SYSTEM StopperingModule (* Module Stoppering, generated from its module specification *)
  (* Standard: 61499-2 *)
  APPLICATION Stoppering (* Module Stoppering on target pc (localhost, IO modbus; generated by modgen) *)
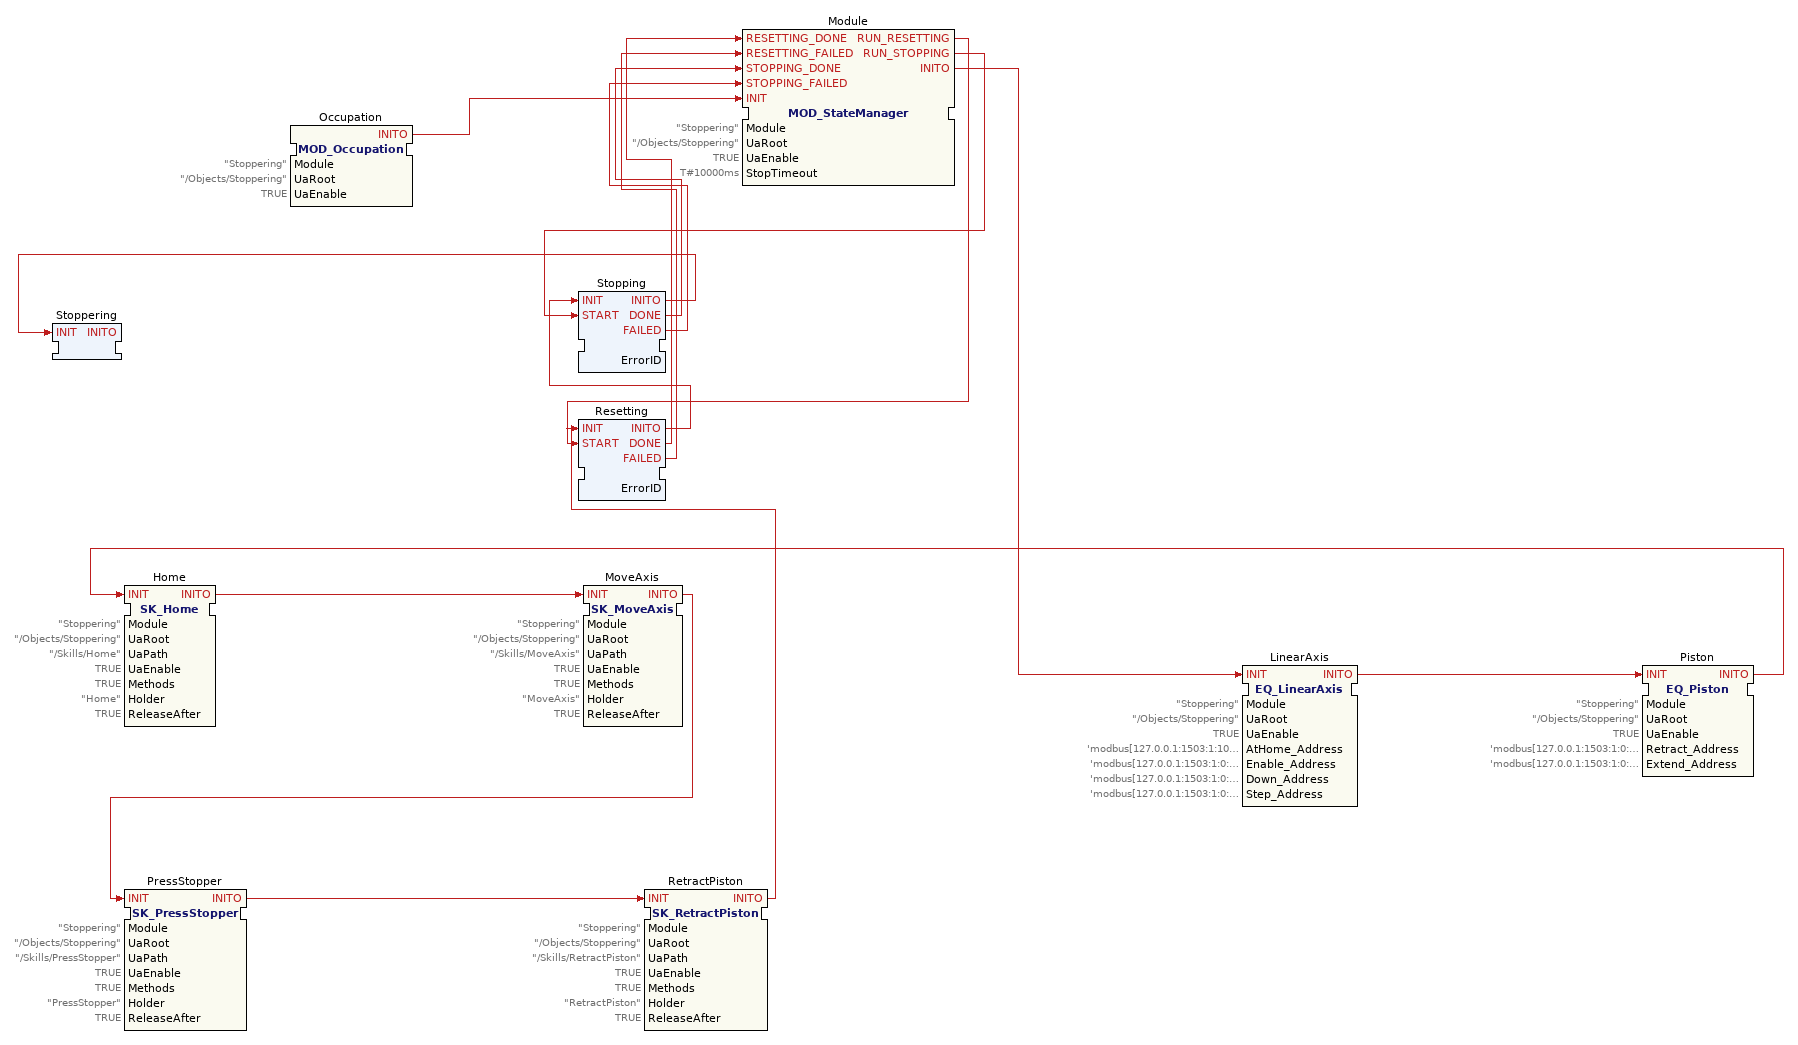
    (* Group ModuleLevel: Module level: occupation, PackML state manager, start-up and the target's IO lines *)
    (* Group ModuleLevelSkills: Module level skills: Control, Sequences (Execute, Stop) of skill primitives and Release; OPC UA /Skills/<name> *)
    (* Group Procedures: Procedures the module state manager runs while Resetting and Stopping *)
    (* Group SkillPrimitives: Skill primitives: one equipment command until a sensor or a time; OPC UA /Skills/<name> *)
    (* Group EquipmentIO: Equipment IO: the only owners of the IO points; skills send them output values over local channels *)
    FBS
      Occupation : modlib::MOD_Occupation(Module := "Stoppering", UaRoot := "/Objects/Stoppering", UaEnable := TRUE); (* Who may command the module. A client calls Occupy(Session) at /Objects/Stoppering/Occupation first; until it calls Release, only commands with that session id are accepted. Every block hears the owner on loc[Stoppering/owner]. *) {SET_ATTRIBUTE(GroupName, ModuleLevel)}
      Module : modlib::MOD_StateManager(Module := "Stoppering", UaRoot := "/Objects/Stoppering", UaEnable := TRUE, StopTimeout := T#10000ms); (* The module's PackML state. The owner calls Reset, Start, Stop, Abort or Clear at /Objects/Stoppering/Module; State is at /Objects/Stoppering/Module/State and on loc[Stoppering/state]. Reset runs the Resetting procedure, Stop the Stopping procedure; skills may be started only in Execute. *) {SET_ATTRIBUTE(GroupName, ModuleLevel)}
      LinearAxis : stoppering::EQ_LinearAxis(Module := "Stoppering", UaRoot := "/Objects/Stoppering", UaEnable := TRUE, AtHome_Address := 'modbus[127.0.0.1:1503:1:10:d0:]', Enable_Address := 'modbus[127.0.0.1:1503:1:0::c0]', Down_Address := 'modbus[127.0.0.1:1503:1:0::c1]', Step_Address := 'modbus[127.0.0.1:1503:1:0::h0]'); (* Equipment LinearAxis: Lift of the stoppering head, a stepper motor through a step and direction driver, with a limit switch at the top (home). The only block that touches its pins (AtHome = modbus[127.0.0.1:1503:1:10:d0:], Enable = modbus[127.0.0.1:1503:1:0::c0], Down = modbus[127.0.0.1:1503:1:0::c1], Step = modbus[127.0.0.1:1503:1:0::h0]). Skills send it what to switch on loc[Stoppering/LinearAxis/cmd]; it reports its inputs on loc[Stoppering/LinearAxis/state] and at /Objects/Stoppering/Equipment/LinearAxis. *) {SET_ATTRIBUTE(GroupName, EquipmentIO)}
      Piston : stoppering::EQ_Piston(Module := "Stoppering", UaRoot := "/Objects/Stoppering", UaEnable := TRUE, Retract_Address := 'modbus[127.0.0.1:1503:1:0::c2]', Extend_Address := 'modbus[127.0.0.1:1503:1:0::c3]'); (* Equipment Piston: Small linear actuator that presses the stopper in, through an L298N (IN1 retract, IN2 extend); no sensors. The only block that touches its pins (Retract = modbus[127.0.0.1:1503:1:0::c2], Extend = modbus[127.0.0.1:1503:1:0::c3]). Skills send it what to switch on loc[Stoppering/Piston/cmd]; it reports its inputs on loc[Stoppering/Piston/state] and at /Objects/Stoppering/Equipment/Piston. *) {SET_ATTRIBUTE(GroupName, EquipmentIO)}
      Home : stoppering::SK_Home(Module := "Stoppering", UaRoot := "/Objects/Stoppering", UaPath := "/Skills/Home", UaEnable := TRUE, Methods := TRUE, Holder := "Home", ReleaseAfter := TRUE); (* Skill Home, offered on its own: Head up to the limit switch; from there its position is known, using LinearAxis. A client calls Start (with the parameters), Stop, Abort or Reset at /Objects/Stoppering/Skills/Home; State, ErrorID, Parameters and Results are there too. *) {SET_ATTRIBUTE(GroupName, SkillPrimitives)}
      MoveAxis : stoppering::SK_MoveAxis(Module := "Stoppering", UaRoot := "/Objects/Stoppering", UaPath := "/Skills/MoveAxis", UaEnable := TRUE, Methods := TRUE, Holder := "MoveAxis", ReleaseAfter := TRUE); (* Skill MoveAxis, offered on its own: Head to Position, measured down from the limit switch; the direction follows from where it is, using LinearAxis. A client calls Start (with the parameters), Stop, Abort or Reset at /Objects/Stoppering/Skills/MoveAxis; State, ErrorID, Parameters and Results are there too. *) {SET_ATTRIBUTE(GroupName, SkillPrimitives)}
      PressStopper : stoppering::SK_PressStopper(Module := "Stoppering", UaRoot := "/Objects/Stoppering", UaPath := "/Skills/PressStopper", UaEnable := TRUE, Methods := TRUE, Holder := "PressStopper", ReleaseAfter := TRUE); (* Skill PressStopper, offered on its own: Press the stopper in, the piston out for the stroke and back in (open loop, by time), using Piston. A client calls Start (with the parameters), Stop, Abort or Reset at /Objects/Stoppering/Skills/PressStopper; State, ErrorID, Parameters and Results are there too. *) {SET_ATTRIBUTE(GroupName, SkillPrimitives)}
      RetractPiston : stoppering::SK_RetractPiston(Module := "Stoppering", UaRoot := "/Objects/Stoppering", UaPath := "/Skills/RetractPiston", UaEnable := TRUE, Methods := TRUE, Holder := "RetractPiston", ReleaseAfter := TRUE); (* Skill RetractPiston, offered on its own: Piston back in for the stroke (open loop); for a piston left out by an abort, using Piston. A client calls Start (with the parameters), Stop, Abort or Reset at /Objects/Stoppering/Skills/RetractPiston; State, ErrorID, Parameters and Results are there too. *) {SET_ATTRIBUTE(GroupName, SkillPrimitives)}
    END_FBS
    SUBAPPLICATION Resetting (* Procedure the module runs while Resetting *)
      {SET_ATTRIBUTE(GroupName, Procedures)}
      EVENT_INPUT
        INIT : EInit;
        START;
      END_EVENT
      EVENT_OUTPUT
        INITO : EInit;
        DONE;
        FAILED;
      END_EVENT
      VAR_OUTPUT
        ErrorID : UINT;
      END_VAR
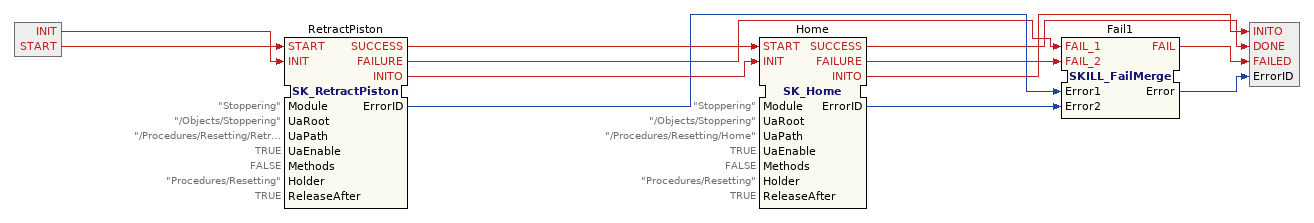
      FBS
        RetractPiston : stoppering::SK_RetractPiston(Module := "Stoppering", UaRoot := "/Objects/Stoppering", UaPath := "/Procedures/Resetting/RetractPiston", UaEnable := TRUE, Methods := FALSE, Holder := "Procedures/Resetting", ReleaseAfter := TRUE); (* Step 1 of Resetting: runs the skill RetractPiston. Its State and ErrorID are at /Objects/Stoppering/Procedures/Resetting/RetractPiston; it keeps the equipment under the name Procedures/Resetting. *)
        Home : stoppering::SK_Home(Module := "Stoppering", UaRoot := "/Objects/Stoppering", UaPath := "/Procedures/Resetting/Home", UaEnable := TRUE, Methods := FALSE, Holder := "Procedures/Resetting", ReleaseAfter := TRUE); (* Step 2 of Resetting: runs the skill Home. Its State and ErrorID are at /Objects/Stoppering/Procedures/Resetting/Home; it keeps the equipment under the name Procedures/Resetting. *)
        Fail1 : modlib::SKILL_FailMerge; (* Joins the failures of the steps into one (with its error code), so any step's failure ends the sequence. *)
      END_FBS
      EVENT_CONNECTIONS
        RetractPiston.SUCCESS TO Home.START;
        START TO RetractPiston.START;
        Home.SUCCESS TO DONE;
        RetractPiston.FAILURE TO Fail1.FAIL_1;
        Home.FAILURE TO Fail1.FAIL_2;
        Fail1.FAIL TO FAILED;
        INIT TO RetractPiston.INIT;
        Home.INITO TO INITO;
        RetractPiston.INITO TO Home.INIT;
      END_CONNECTIONS
      DATA_CONNECTIONS
        RetractPiston.ErrorID TO Fail1.Error1;
        Home.ErrorID TO Fail1.Error2;
        Fail1.Error TO ErrorID;
      END_CONNECTIONS
    END_SUBAPPLICATION
    SUBAPPLICATION Stopping (* Procedure the module runs while Stopping *)
      {SET_ATTRIBUTE(GroupName, Procedures)}
      EVENT_INPUT
        INIT : EInit;
        START;
      END_EVENT
      EVENT_OUTPUT
        INITO : EInit;
        DONE;
        FAILED;
      END_EVENT
      VAR_OUTPUT
        ErrorID : UINT;
      END_VAR
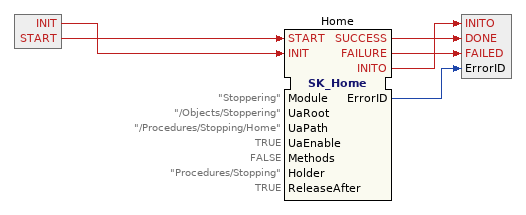
      FBS
        Home : stoppering::SK_Home(Module := "Stoppering", UaRoot := "/Objects/Stoppering", UaPath := "/Procedures/Stopping/Home", UaEnable := TRUE, Methods := FALSE, Holder := "Procedures/Stopping", ReleaseAfter := TRUE); (* Step 1 of Stopping: runs the skill Home. Its State and ErrorID are at /Objects/Stoppering/Procedures/Stopping/Home; it keeps the equipment under the name Procedures/Stopping. *)
      END_FBS
      EVENT_CONNECTIONS
        START TO Home.START;
        Home.SUCCESS TO DONE;
        Home.FAILURE TO FAILED;
        INIT TO Home.INIT;
        Home.INITO TO INITO;
      END_CONNECTIONS
      DATA_CONNECTIONS
        Home.ErrorID TO ErrorID;
      END_CONNECTIONS
    END_SUBAPPLICATION
    SUBAPPLICATION Stoppering (* Module level skill Stoppering: Head down onto the vial, press the stopper in, head up again *)
      {SET_ATTRIBUTE(GroupName, ModuleLevelSkills)}
      EVENT_INPUT
        INIT : EInit;
      END_EVENT
      EVENT_OUTPUT
        INITO : EInit;
      END_EVENT
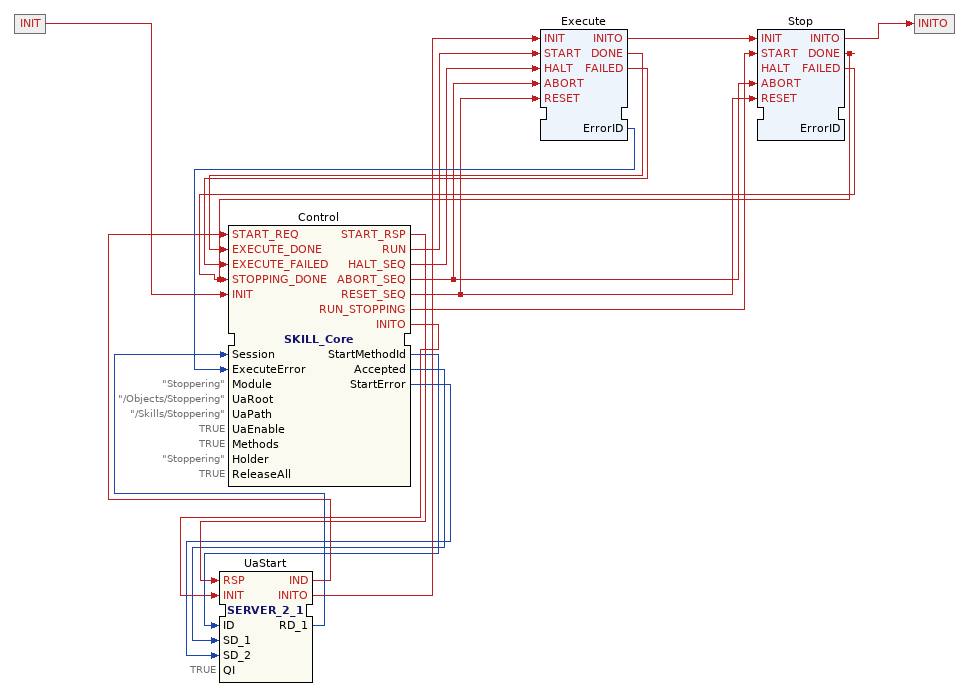
      (* Group Core: The skill's state machine: Stop, Abort, Reset, State and ErrorID over OPC UA; gives up everything the skill holds when a run ends *)
      (* Group Start: The Start method: one block per parameter (range check, value for this run), the values published *)
      (* Group Sequences: What the skill does: Execute, and Stop when it is interrupted; private skill primitives in order *)
      FBS
        Control : modlib::SKILL_Core(Module := "Stoppering", UaRoot := "/Objects/Stoppering", UaPath := "/Skills/Stoppering", UaEnable := TRUE, Methods := TRUE, Holder := "Stoppering", ReleaseAll := TRUE); (* The state machine of the skill Stoppering: checks a client's Start (occupation, module in Execute, not running, values in range), publishes State and ErrorID at /Objects/Stoppering/Skills/Stoppering, offers Stop, Abort and Reset there, starts Execute and runs Stop when the skill is stopped. *) {SET_ATTRIBUTE(GroupName, Core)}
        UaStart : iec61499::net::SERVER_2_1(QI := TRUE); (* The OPC UA method Start of Stoppering: a client's call (session id and parameters) arrives here; the parameters are checked, then Control answers Accepted or an error code. *) {SET_ATTRIBUTE(GroupName, Start)}
      END_FBS
      SUBAPPLICATION Execute (* Stoppering: execute sequence *)
        {SET_ATTRIBUTE(GroupName, Sequences)}
        EVENT_INPUT
          INIT : EInit;
          START;
          HALT;
          ABORT;
          RESET;
        END_EVENT
        EVENT_OUTPUT
          INITO : EInit;
          DONE;
          FAILED;
        END_EVENT
        VAR_OUTPUT
          ErrorID : UINT;
        END_VAR
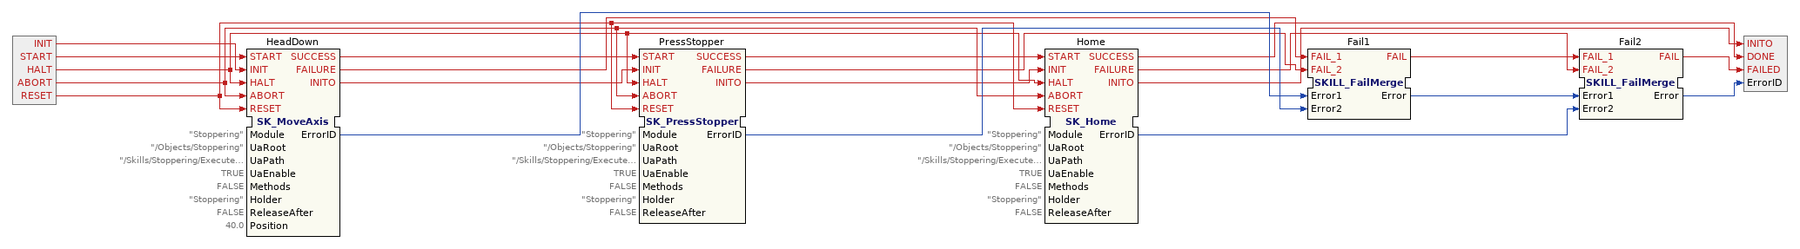
        FBS
          HeadDown : stoppering::SK_MoveAxis(Module := "Stoppering", UaRoot := "/Objects/Stoppering", UaPath := "/Skills/Stoppering/Execute/HeadDown", UaEnable := TRUE, Methods := FALSE, Holder := "Stoppering", ReleaseAfter := FALSE, Position := 40.0); (* Step 1 of Stoppering / Execute: runs the skill MoveAxis with Position = 40.0. Its State and ErrorID are at /Objects/Stoppering/Skills/Stoppering/Execute/HeadDown; it keeps the equipment under the name Stoppering. *)
          PressStopper : stoppering::SK_PressStopper(Module := "Stoppering", UaRoot := "/Objects/Stoppering", UaPath := "/Skills/Stoppering/Execute/PressStopper", UaEnable := TRUE, Methods := FALSE, Holder := "Stoppering", ReleaseAfter := FALSE); (* Step 2 of Stoppering / Execute: runs the skill PressStopper. Its State and ErrorID are at /Objects/Stoppering/Skills/Stoppering/Execute/PressStopper; it keeps the equipment under the name Stoppering. *)
          Home : stoppering::SK_Home(Module := "Stoppering", UaRoot := "/Objects/Stoppering", UaPath := "/Skills/Stoppering/Execute/Home", UaEnable := TRUE, Methods := FALSE, Holder := "Stoppering", ReleaseAfter := FALSE); (* Step 3 of Stoppering / Execute: runs the skill Home. Its State and ErrorID are at /Objects/Stoppering/Skills/Stoppering/Execute/Home; it keeps the equipment under the name Stoppering. *)
          Fail1 : modlib::SKILL_FailMerge; (* Joins the failures of the steps into one (with its error code), so any step's failure ends the sequence. *)
          Fail2 : modlib::SKILL_FailMerge; (* Joins the failures of the steps into one (with its error code), so any step's failure ends the sequence. *)
        END_FBS
        EVENT_CONNECTIONS
          HeadDown.SUCCESS TO PressStopper.START;
          PressStopper.SUCCESS TO Home.START;
          START TO HeadDown.START;
          Home.SUCCESS TO DONE;
          HeadDown.FAILURE TO Fail1.FAIL_1;
          PressStopper.FAILURE TO Fail1.FAIL_2;
          Fail1.FAIL TO Fail2.FAIL_1;
          Home.FAILURE TO Fail2.FAIL_2;
          Fail2.FAIL TO FAILED;
          INIT TO HeadDown.INIT;
          Home.INITO TO INITO;
          HeadDown.INITO TO PressStopper.INIT;
          PressStopper.INITO TO Home.INIT;
          HALT TO HeadDown.HALT;
          HALT TO PressStopper.HALT;
          HALT TO Home.HALT;
          ABORT TO HeadDown.ABORT;
          ABORT TO PressStopper.ABORT;
          ABORT TO Home.ABORT;
          RESET TO HeadDown.RESET;
          RESET TO PressStopper.RESET;
          RESET TO Home.RESET;
        END_CONNECTIONS
        DATA_CONNECTIONS
          HeadDown.ErrorID TO Fail1.Error1;
          PressStopper.ErrorID TO Fail1.Error2;
          Fail1.Error TO Fail2.Error1;
          Home.ErrorID TO Fail2.Error2;
          Fail2.Error TO ErrorID;
        END_CONNECTIONS
      END_SUBAPPLICATION
      SUBAPPLICATION Stop (* Stoppering: stop sequence *)
        {SET_ATTRIBUTE(GroupName, Sequences)}
        EVENT_INPUT
          INIT : EInit;
          START;
          HALT;
          ABORT;
          RESET;
        END_EVENT
        EVENT_OUTPUT
          INITO : EInit;
          DONE;
          FAILED;
        END_EVENT
        VAR_OUTPUT
          ErrorID : UINT;
        END_VAR
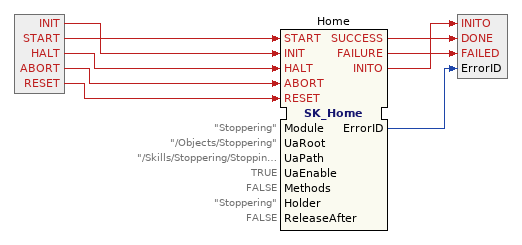
        FBS
          Home : stoppering::SK_Home(Module := "Stoppering", UaRoot := "/Objects/Stoppering", UaPath := "/Skills/Stoppering/Stopping/Home", UaEnable := TRUE, Methods := FALSE, Holder := "Stoppering", ReleaseAfter := FALSE); (* Step 1 of Stoppering / Stop: runs the skill Home. Its State and ErrorID are at /Objects/Stoppering/Skills/Stoppering/Stopping/Home; it keeps the equipment under the name Stoppering. *)
        END_FBS
        EVENT_CONNECTIONS
          START TO Home.START;
          Home.SUCCESS TO DONE;
          Home.FAILURE TO FAILED;
          INIT TO Home.INIT;
          Home.INITO TO INITO;
          HALT TO Home.HALT;
          ABORT TO Home.ABORT;
          RESET TO Home.RESET;
        END_CONNECTIONS
        DATA_CONNECTIONS
          Home.ErrorID TO ErrorID;
        END_CONNECTIONS
      END_SUBAPPLICATION
      EVENT_CONNECTIONS
        Control.START_RSP TO UaStart.RSP;
        UaStart.IND TO Control.START_REQ;
        Control.RUN TO Execute.START;
        Control.HALT_SEQ TO Execute.HALT;
        Control.ABORT_SEQ TO Execute.ABORT;
        Control.RESET_SEQ TO Execute.RESET;
        Execute.DONE TO Control.EXECUTE_DONE;
        Execute.FAILED TO Control.EXECUTE_FAILED;
        Control.RUN_STOPPING TO Stop.START;
        Control.ABORT_SEQ TO Stop.ABORT;
        Control.RESET_SEQ TO Stop.RESET;
        Stop.DONE TO Control.STOPPING_DONE;
        Stop.FAILED TO Control.STOPPING_DONE;
        INIT TO Control.INIT;
        Control.INITO TO UaStart.INIT;
        UaStart.INITO TO Execute.INIT;
        Execute.INITO TO Stop.INIT;
        Stop.INITO TO INITO;
      END_CONNECTIONS
      DATA_CONNECTIONS
        Control.StartMethodId TO UaStart.ID;
        UaStart.RD_1 TO Control.Session;
        Control.Accepted TO UaStart.SD_1;
        Control.StartError TO UaStart.SD_2;
        Execute.ErrorID TO Control.ExecuteError;
      END_CONNECTIONS
    END_SUBAPPLICATION
    EVENT_CONNECTIONS
      Module.RUN_RESETTING TO Resetting.START;
      Resetting.DONE TO Module.RESETTING_DONE;
      Resetting.FAILED TO Module.RESETTING_FAILED;
      Module.RUN_STOPPING TO Stopping.START;
      Stopping.DONE TO Module.STOPPING_DONE;
      Stopping.FAILED TO Module.STOPPING_FAILED;
      Occupation.INITO TO Module.INIT;
      Module.INITO TO LinearAxis.INIT;
      LinearAxis.INITO TO Piston.INIT;
      Piston.INITO TO Home.INIT;
      Home.INITO TO MoveAxis.INIT;
      MoveAxis.INITO TO PressStopper.INIT;
      PressStopper.INITO TO RetractPiston.INIT;
      RetractPiston.INITO TO Resetting.INIT;
      Resetting.INITO TO Stopping.INIT;
      Stopping.INITO TO Stoppering.INIT;
    END_CONNECTIONS
  END_APPLICATION
  APPLICATION Stoppering_pi (* Module Stoppering on target pi (192.168.0.134, IO gpio; generated by modgen) *)
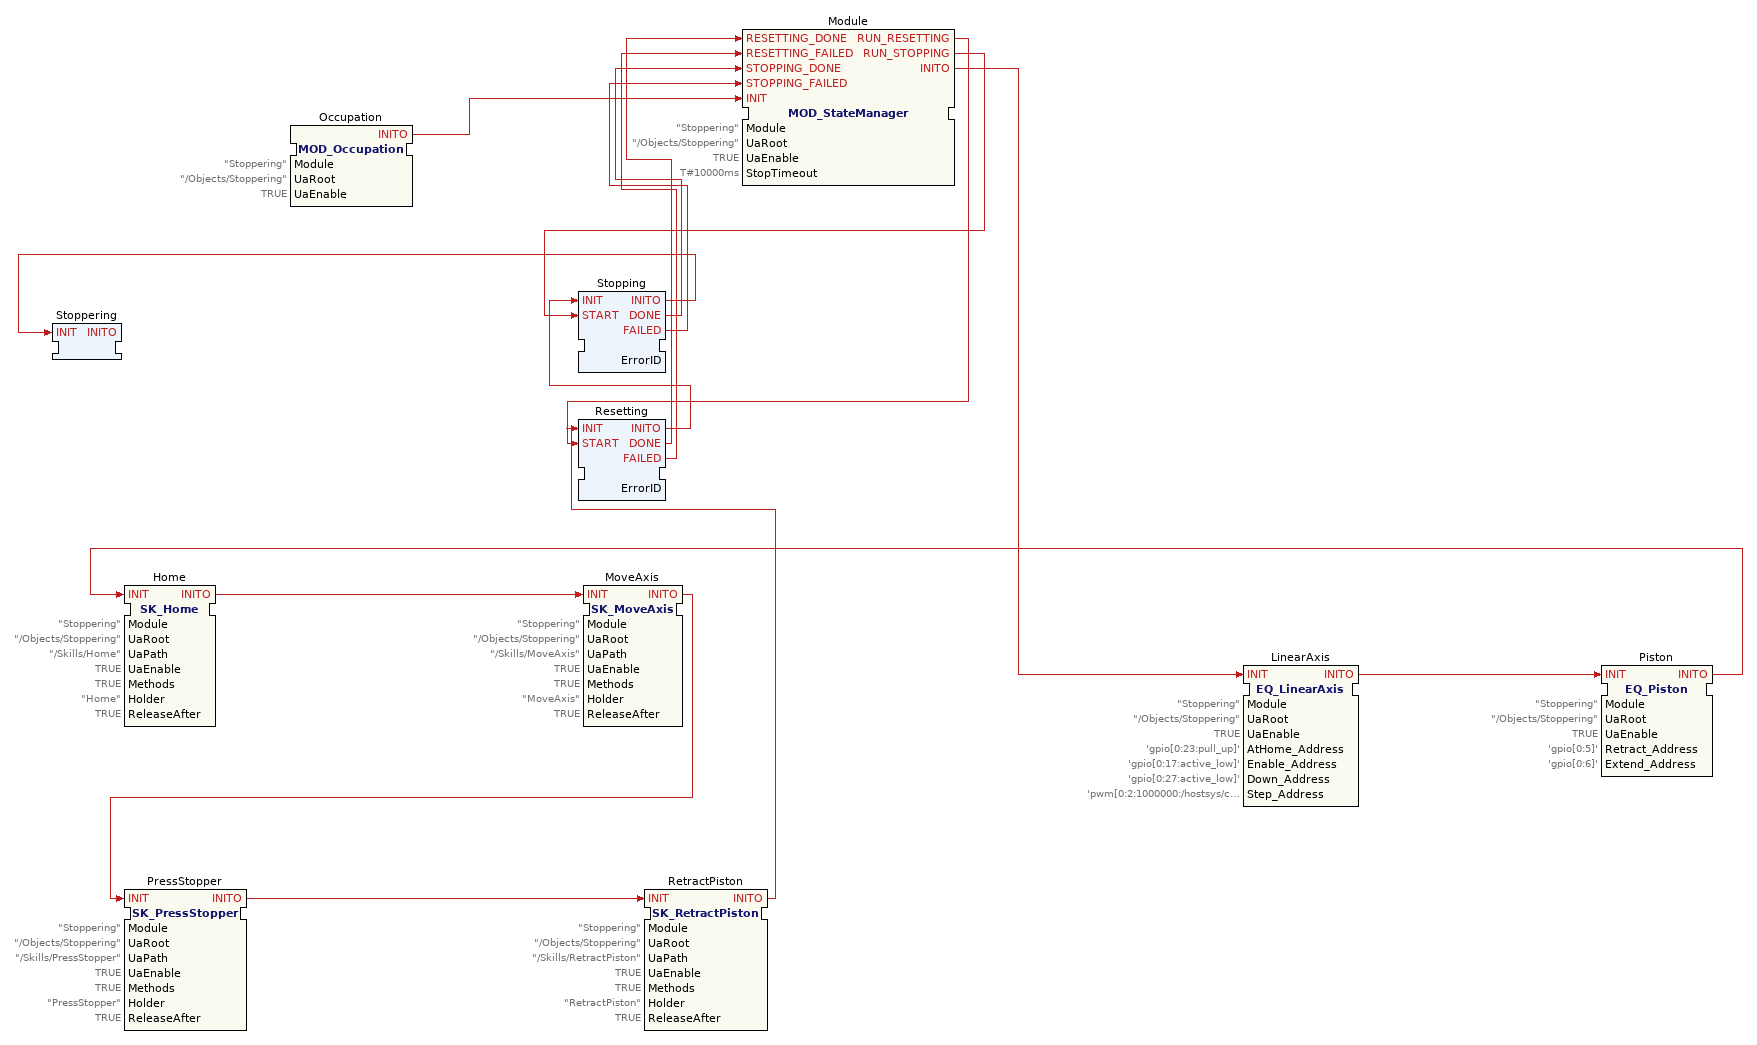
    (* Group ModuleLevel: Module level: occupation, PackML state manager, start-up and the target's IO lines *)
    (* Group ModuleLevelSkills: Module level skills: Control, Sequences (Execute, Stop) of skill primitives and Release; OPC UA /Skills/<name> *)
    (* Group Procedures: Procedures the module state manager runs while Resetting and Stopping *)
    (* Group SkillPrimitives: Skill primitives: one equipment command until a sensor or a time; OPC UA /Skills/<name> *)
    (* Group EquipmentIO: Equipment IO: the only owners of the IO points; skills send them output values over local channels *)
    FBS
      Occupation : modlib::MOD_Occupation(Module := "Stoppering", UaRoot := "/Objects/Stoppering", UaEnable := TRUE); (* Who may command the module. A client calls Occupy(Session) at /Objects/Stoppering/Occupation first; until it calls Release, only commands with that session id are accepted. Every block hears the owner on loc[Stoppering/owner]. *) {SET_ATTRIBUTE(GroupName, ModuleLevel)}
      Module : modlib::MOD_StateManager(Module := "Stoppering", UaRoot := "/Objects/Stoppering", UaEnable := TRUE, StopTimeout := T#10000ms); (* The module's PackML state. The owner calls Reset, Start, Stop, Abort or Clear at /Objects/Stoppering/Module; State is at /Objects/Stoppering/Module/State and on loc[Stoppering/state]. Reset runs the Resetting procedure, Stop the Stopping procedure; skills may be started only in Execute. *) {SET_ATTRIBUTE(GroupName, ModuleLevel)}
      LinearAxis : stoppering::EQ_LinearAxis(Module := "Stoppering", UaRoot := "/Objects/Stoppering", UaEnable := TRUE, AtHome_Address := 'gpio[0:23:pull_up]', Enable_Address := 'gpio[0:17:active_low]', Down_Address := 'gpio[0:27:active_low]', Step_Address := 'pwm[0:2:1000000:/hostsys/class/pwm]'); (* Equipment LinearAxis: Lift of the stoppering head, a stepper motor through a step and direction driver, with a limit switch at the top (home). The only block that touches its pins (AtHome = gpio[0:23:pull_up], Enable = gpio[0:17:active_low], Down = gpio[0:27:active_low], Step = pwm[0:2:1000000:/hostsys/class/pwm]). Skills send it what to switch on loc[Stoppering/LinearAxis/cmd]; it reports its inputs on loc[Stoppering/LinearAxis/state] and at /Objects/Stoppering/Equipment/LinearAxis. *) {SET_ATTRIBUTE(GroupName, EquipmentIO)}
      Piston : stoppering::EQ_Piston(Module := "Stoppering", UaRoot := "/Objects/Stoppering", UaEnable := TRUE, Retract_Address := 'gpio[0:5]', Extend_Address := 'gpio[0:6]'); (* Equipment Piston: Small linear actuator that presses the stopper in, through an L298N (IN1 retract, IN2 extend); no sensors. The only block that touches its pins (Retract = gpio[0:5], Extend = gpio[0:6]). Skills send it what to switch on loc[Stoppering/Piston/cmd]; it reports its inputs on loc[Stoppering/Piston/state] and at /Objects/Stoppering/Equipment/Piston. *) {SET_ATTRIBUTE(GroupName, EquipmentIO)}
      Home : stoppering::SK_Home(Module := "Stoppering", UaRoot := "/Objects/Stoppering", UaPath := "/Skills/Home", UaEnable := TRUE, Methods := TRUE, Holder := "Home", ReleaseAfter := TRUE); (* Skill Home, offered on its own: Head up to the limit switch; from there its position is known, using LinearAxis. A client calls Start (with the parameters), Stop, Abort or Reset at /Objects/Stoppering/Skills/Home; State, ErrorID, Parameters and Results are there too. *) {SET_ATTRIBUTE(GroupName, SkillPrimitives)}
      MoveAxis : stoppering::SK_MoveAxis(Module := "Stoppering", UaRoot := "/Objects/Stoppering", UaPath := "/Skills/MoveAxis", UaEnable := TRUE, Methods := TRUE, Holder := "MoveAxis", ReleaseAfter := TRUE); (* Skill MoveAxis, offered on its own: Head to Position, measured down from the limit switch; the direction follows from where it is, using LinearAxis. A client calls Start (with the parameters), Stop, Abort or Reset at /Objects/Stoppering/Skills/MoveAxis; State, ErrorID, Parameters and Results are there too. *) {SET_ATTRIBUTE(GroupName, SkillPrimitives)}
      PressStopper : stoppering::SK_PressStopper(Module := "Stoppering", UaRoot := "/Objects/Stoppering", UaPath := "/Skills/PressStopper", UaEnable := TRUE, Methods := TRUE, Holder := "PressStopper", ReleaseAfter := TRUE); (* Skill PressStopper, offered on its own: Press the stopper in, the piston out for the stroke and back in (open loop, by time), using Piston. A client calls Start (with the parameters), Stop, Abort or Reset at /Objects/Stoppering/Skills/PressStopper; State, ErrorID, Parameters and Results are there too. *) {SET_ATTRIBUTE(GroupName, SkillPrimitives)}
      RetractPiston : stoppering::SK_RetractPiston(Module := "Stoppering", UaRoot := "/Objects/Stoppering", UaPath := "/Skills/RetractPiston", UaEnable := TRUE, Methods := TRUE, Holder := "RetractPiston", ReleaseAfter := TRUE); (* Skill RetractPiston, offered on its own: Piston back in for the stroke (open loop); for a piston left out by an abort, using Piston. A client calls Start (with the parameters), Stop, Abort or Reset at /Objects/Stoppering/Skills/RetractPiston; State, ErrorID, Parameters and Results are there too. *) {SET_ATTRIBUTE(GroupName, SkillPrimitives)}
    END_FBS
    SUBAPPLICATION Resetting (* Procedure the module runs while Resetting *)
      {SET_ATTRIBUTE(GroupName, Procedures)}
      EVENT_INPUT
        INIT : EInit;
        START;
      END_EVENT
      EVENT_OUTPUT
        INITO : EInit;
        DONE;
        FAILED;
      END_EVENT
      VAR_OUTPUT
        ErrorID : UINT;
      END_VAR
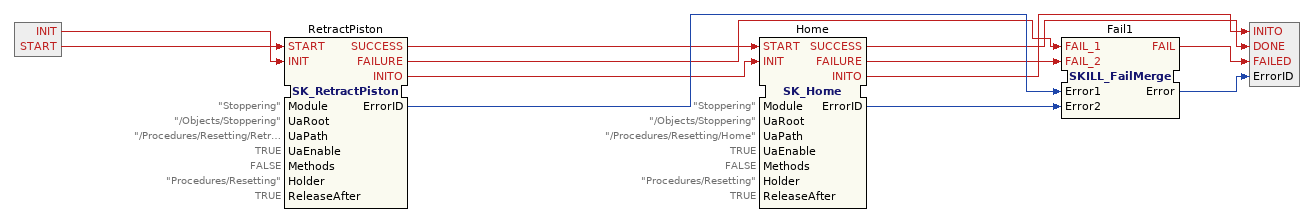
      FBS
        RetractPiston : stoppering::SK_RetractPiston(Module := "Stoppering", UaRoot := "/Objects/Stoppering", UaPath := "/Procedures/Resetting/RetractPiston", UaEnable := TRUE, Methods := FALSE, Holder := "Procedures/Resetting", ReleaseAfter := TRUE); (* Step 1 of Resetting: runs the skill RetractPiston. Its State and ErrorID are at /Objects/Stoppering/Procedures/Resetting/RetractPiston; it keeps the equipment under the name Procedures/Resetting. *)
        Home : stoppering::SK_Home(Module := "Stoppering", UaRoot := "/Objects/Stoppering", UaPath := "/Procedures/Resetting/Home", UaEnable := TRUE, Methods := FALSE, Holder := "Procedures/Resetting", ReleaseAfter := TRUE); (* Step 2 of Resetting: runs the skill Home. Its State and ErrorID are at /Objects/Stoppering/Procedures/Resetting/Home; it keeps the equipment under the name Procedures/Resetting. *)
        Fail1 : modlib::SKILL_FailMerge; (* Joins the failures of the steps into one (with its error code), so any step's failure ends the sequence. *)
      END_FBS
      EVENT_CONNECTIONS
        RetractPiston.SUCCESS TO Home.START;
        START TO RetractPiston.START;
        Home.SUCCESS TO DONE;
        RetractPiston.FAILURE TO Fail1.FAIL_1;
        Home.FAILURE TO Fail1.FAIL_2;
        Fail1.FAIL TO FAILED;
        INIT TO RetractPiston.INIT;
        Home.INITO TO INITO;
        RetractPiston.INITO TO Home.INIT;
      END_CONNECTIONS
      DATA_CONNECTIONS
        RetractPiston.ErrorID TO Fail1.Error1;
        Home.ErrorID TO Fail1.Error2;
        Fail1.Error TO ErrorID;
      END_CONNECTIONS
    END_SUBAPPLICATION
    SUBAPPLICATION Stopping (* Procedure the module runs while Stopping *)
      {SET_ATTRIBUTE(GroupName, Procedures)}
      EVENT_INPUT
        INIT : EInit;
        START;
      END_EVENT
      EVENT_OUTPUT
        INITO : EInit;
        DONE;
        FAILED;
      END_EVENT
      VAR_OUTPUT
        ErrorID : UINT;
      END_VAR
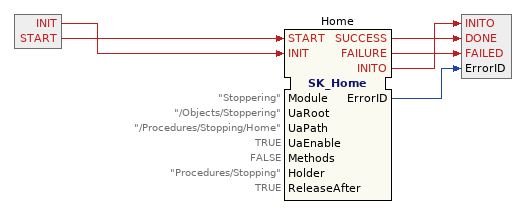
      FBS
        Home : stoppering::SK_Home(Module := "Stoppering", UaRoot := "/Objects/Stoppering", UaPath := "/Procedures/Stopping/Home", UaEnable := TRUE, Methods := FALSE, Holder := "Procedures/Stopping", ReleaseAfter := TRUE); (* Step 1 of Stopping: runs the skill Home. Its State and ErrorID are at /Objects/Stoppering/Procedures/Stopping/Home; it keeps the equipment under the name Procedures/Stopping. *)
      END_FBS
      EVENT_CONNECTIONS
        START TO Home.START;
        Home.SUCCESS TO DONE;
        Home.FAILURE TO FAILED;
        INIT TO Home.INIT;
        Home.INITO TO INITO;
      END_CONNECTIONS
      DATA_CONNECTIONS
        Home.ErrorID TO ErrorID;
      END_CONNECTIONS
    END_SUBAPPLICATION
    SUBAPPLICATION Stoppering (* Module level skill Stoppering: Head down onto the vial, press the stopper in, head up again *)
      {SET_ATTRIBUTE(GroupName, ModuleLevelSkills)}
      EVENT_INPUT
        INIT : EInit;
      END_EVENT
      EVENT_OUTPUT
        INITO : EInit;
      END_EVENT
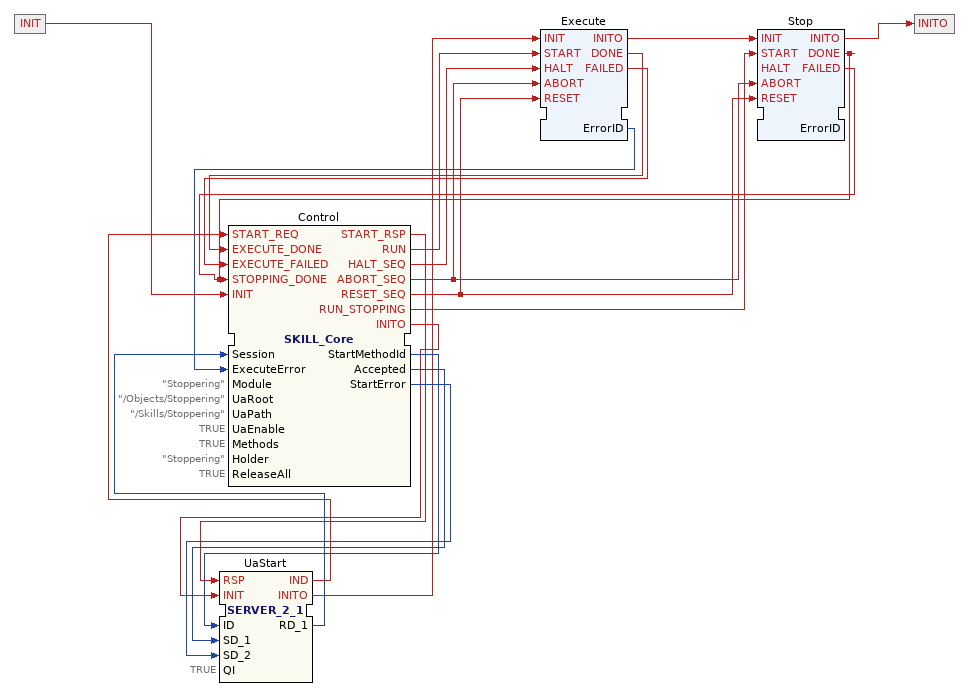
      (* Group Core: The skill's state machine: Stop, Abort, Reset, State and ErrorID over OPC UA; gives up everything the skill holds when a run ends *)
      (* Group Start: The Start method: one block per parameter (range check, value for this run), the values published *)
      (* Group Sequences: What the skill does: Execute, and Stop when it is interrupted; private skill primitives in order *)
      FBS
        Control : modlib::SKILL_Core(Module := "Stoppering", UaRoot := "/Objects/Stoppering", UaPath := "/Skills/Stoppering", UaEnable := TRUE, Methods := TRUE, Holder := "Stoppering", ReleaseAll := TRUE); (* The state machine of the skill Stoppering: checks a client's Start (occupation, module in Execute, not running, values in range), publishes State and ErrorID at /Objects/Stoppering/Skills/Stoppering, offers Stop, Abort and Reset there, starts Execute and runs Stop when the skill is stopped. *) {SET_ATTRIBUTE(GroupName, Core)}
        UaStart : iec61499::net::SERVER_2_1(QI := TRUE); (* The OPC UA method Start of Stoppering: a client's call (session id and parameters) arrives here; the parameters are checked, then Control answers Accepted or an error code. *) {SET_ATTRIBUTE(GroupName, Start)}
      END_FBS
      SUBAPPLICATION Execute (* Stoppering: execute sequence *)
        {SET_ATTRIBUTE(GroupName, Sequences)}
        EVENT_INPUT
          INIT : EInit;
          START;
          HALT;
          ABORT;
          RESET;
        END_EVENT
        EVENT_OUTPUT
          INITO : EInit;
          DONE;
          FAILED;
        END_EVENT
        VAR_OUTPUT
          ErrorID : UINT;
        END_VAR
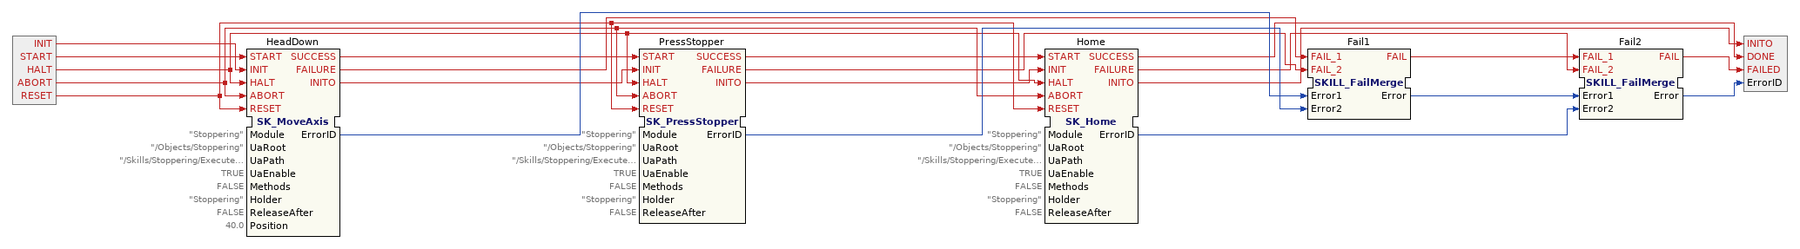
        FBS
          HeadDown : stoppering::SK_MoveAxis(Module := "Stoppering", UaRoot := "/Objects/Stoppering", UaPath := "/Skills/Stoppering/Execute/HeadDown", UaEnable := TRUE, Methods := FALSE, Holder := "Stoppering", ReleaseAfter := FALSE, Position := 40.0); (* Step 1 of Stoppering / Execute: runs the skill MoveAxis with Position = 40.0. Its State and ErrorID are at /Objects/Stoppering/Skills/Stoppering/Execute/HeadDown; it keeps the equipment under the name Stoppering. *)
          PressStopper : stoppering::SK_PressStopper(Module := "Stoppering", UaRoot := "/Objects/Stoppering", UaPath := "/Skills/Stoppering/Execute/PressStopper", UaEnable := TRUE, Methods := FALSE, Holder := "Stoppering", ReleaseAfter := FALSE); (* Step 2 of Stoppering / Execute: runs the skill PressStopper. Its State and ErrorID are at /Objects/Stoppering/Skills/Stoppering/Execute/PressStopper; it keeps the equipment under the name Stoppering. *)
          Home : stoppering::SK_Home(Module := "Stoppering", UaRoot := "/Objects/Stoppering", UaPath := "/Skills/Stoppering/Execute/Home", UaEnable := TRUE, Methods := FALSE, Holder := "Stoppering", ReleaseAfter := FALSE); (* Step 3 of Stoppering / Execute: runs the skill Home. Its State and ErrorID are at /Objects/Stoppering/Skills/Stoppering/Execute/Home; it keeps the equipment under the name Stoppering. *)
          Fail1 : modlib::SKILL_FailMerge; (* Joins the failures of the steps into one (with its error code), so any step's failure ends the sequence. *)
          Fail2 : modlib::SKILL_FailMerge; (* Joins the failures of the steps into one (with its error code), so any step's failure ends the sequence. *)
        END_FBS
        EVENT_CONNECTIONS
          HeadDown.SUCCESS TO PressStopper.START;
          PressStopper.SUCCESS TO Home.START;
          START TO HeadDown.START;
          Home.SUCCESS TO DONE;
          HeadDown.FAILURE TO Fail1.FAIL_1;
          PressStopper.FAILURE TO Fail1.FAIL_2;
          Fail1.FAIL TO Fail2.FAIL_1;
          Home.FAILURE TO Fail2.FAIL_2;
          Fail2.FAIL TO FAILED;
          INIT TO HeadDown.INIT;
          Home.INITO TO INITO;
          HeadDown.INITO TO PressStopper.INIT;
          PressStopper.INITO TO Home.INIT;
          HALT TO HeadDown.HALT;
          HALT TO PressStopper.HALT;
          HALT TO Home.HALT;
          ABORT TO HeadDown.ABORT;
          ABORT TO PressStopper.ABORT;
          ABORT TO Home.ABORT;
          RESET TO HeadDown.RESET;
          RESET TO PressStopper.RESET;
          RESET TO Home.RESET;
        END_CONNECTIONS
        DATA_CONNECTIONS
          HeadDown.ErrorID TO Fail1.Error1;
          PressStopper.ErrorID TO Fail1.Error2;
          Fail1.Error TO Fail2.Error1;
          Home.ErrorID TO Fail2.Error2;
          Fail2.Error TO ErrorID;
        END_CONNECTIONS
      END_SUBAPPLICATION
      SUBAPPLICATION Stop (* Stoppering: stop sequence *)
        {SET_ATTRIBUTE(GroupName, Sequences)}
        EVENT_INPUT
          INIT : EInit;
          START;
          HALT;
          ABORT;
          RESET;
        END_EVENT
        EVENT_OUTPUT
          INITO : EInit;
          DONE;
          FAILED;
        END_EVENT
        VAR_OUTPUT
          ErrorID : UINT;
        END_VAR
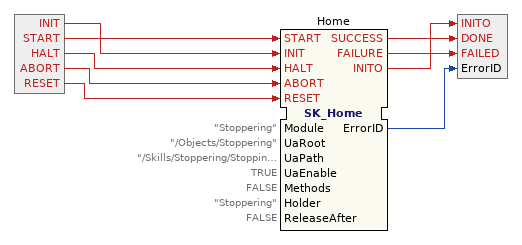
        FBS
          Home : stoppering::SK_Home(Module := "Stoppering", UaRoot := "/Objects/Stoppering", UaPath := "/Skills/Stoppering/Stopping/Home", UaEnable := TRUE, Methods := FALSE, Holder := "Stoppering", ReleaseAfter := FALSE); (* Step 1 of Stoppering / Stop: runs the skill Home. Its State and ErrorID are at /Objects/Stoppering/Skills/Stoppering/Stopping/Home; it keeps the equipment under the name Stoppering. *)
        END_FBS
        EVENT_CONNECTIONS
          START TO Home.START;
          Home.SUCCESS TO DONE;
          Home.FAILURE TO FAILED;
          INIT TO Home.INIT;
          Home.INITO TO INITO;
          HALT TO Home.HALT;
          ABORT TO Home.ABORT;
          RESET TO Home.RESET;
        END_CONNECTIONS
        DATA_CONNECTIONS
          Home.ErrorID TO ErrorID;
        END_CONNECTIONS
      END_SUBAPPLICATION
      EVENT_CONNECTIONS
        Control.START_RSP TO UaStart.RSP;
        UaStart.IND TO Control.START_REQ;
        Control.RUN TO Execute.START;
        Control.HALT_SEQ TO Execute.HALT;
        Control.ABORT_SEQ TO Execute.ABORT;
        Control.RESET_SEQ TO Execute.RESET;
        Execute.DONE TO Control.EXECUTE_DONE;
        Execute.FAILED TO Control.EXECUTE_FAILED;
        Control.RUN_STOPPING TO Stop.START;
        Control.ABORT_SEQ TO Stop.ABORT;
        Control.RESET_SEQ TO Stop.RESET;
        Stop.DONE TO Control.STOPPING_DONE;
        Stop.FAILED TO Control.STOPPING_DONE;
        INIT TO Control.INIT;
        Control.INITO TO UaStart.INIT;
        UaStart.INITO TO Execute.INIT;
        Execute.INITO TO Stop.INIT;
        Stop.INITO TO INITO;
      END_CONNECTIONS
      DATA_CONNECTIONS
        Control.StartMethodId TO UaStart.ID;
        UaStart.RD_1 TO Control.Session;
        Control.Accepted TO UaStart.SD_1;
        Control.StartError TO UaStart.SD_2;
        Execute.ErrorID TO Control.ExecuteError;
      END_CONNECTIONS
    END_SUBAPPLICATION
    EVENT_CONNECTIONS
      Module.RUN_RESETTING TO Resetting.START;
      Resetting.DONE TO Module.RESETTING_DONE;
      Resetting.FAILED TO Module.RESETTING_FAILED;
      Module.RUN_STOPPING TO Stopping.START;
      Stopping.DONE TO Module.STOPPING_DONE;
      Stopping.FAILED TO Module.STOPPING_FAILED;
      Occupation.INITO TO Module.INIT;
      Module.INITO TO LinearAxis.INIT;
      LinearAxis.INITO TO Piston.INIT;
      Piston.INITO TO Home.INIT;
      Home.INITO TO MoveAxis.INIT;
      MoveAxis.INITO TO PressStopper.INIT;
      PressStopper.INITO TO RetractPiston.INIT;
      RetractPiston.INITO TO Resetting.INIT;
      Resetting.INITO TO Stopping.INIT;
      Stopping.INITO TO Stoppering.INIT;
    END_CONNECTIONS
  END_APPLICATION
  DEVICE FORTE_PC : iec61499::system::FORTE_PC(MGR_ID := "localhost:61499" (* Device manager socket ID *))
    {SET_ATTRIBUTE(Profile, HOLOBLOC)}
    RESOURCE RES : iec61499::system::EMB_RES
      EVENT_CONNECTIONS
        START.COLD TO Stoppering.Occupation.INIT;
        START.WARM TO Stoppering.Occupation.INIT;
      END_CONNECTIONS
    END_RESOURCE
  END_DEVICE
  DEVICE FORTE_PI : iec61499::system::FORTE_PC(MGR_ID := "192.168.0.134:61499" (* Device manager socket ID *))
    {SET_ATTRIBUTE(Profile, HOLOBLOC)}
    RESOURCE RES : iec61499::system::EMB_RES
      EVENT_CONNECTIONS
        START.COLD TO Stoppering_pi.Occupation.INIT;
        START.WARM TO Stoppering_pi.Occupation.INIT;
      END_CONNECTIONS
    END_RESOURCE
  END_DEVICE
  MAPPINGS
    Stoppering.Occupation ON FORTE_PC.RES;
    Stoppering.Module ON FORTE_PC.RES;
    Stoppering.LinearAxis ON FORTE_PC.RES;
    Stoppering.Piston ON FORTE_PC.RES;
    Stoppering.Home ON FORTE_PC.RES;
    Stoppering.MoveAxis ON FORTE_PC.RES;
    Stoppering.PressStopper ON FORTE_PC.RES;
    Stoppering.RetractPiston ON FORTE_PC.RES;
    Stoppering.Resetting ON FORTE_PC.RES;
    Stoppering.Stopping ON FORTE_PC.RES;
    Stoppering.Stoppering ON FORTE_PC.RES;
    Stoppering_pi.Occupation ON FORTE_PI.RES;
    Stoppering_pi.Module ON FORTE_PI.RES;
    Stoppering_pi.LinearAxis ON FORTE_PI.RES;
    Stoppering_pi.Piston ON FORTE_PI.RES;
    Stoppering_pi.Home ON FORTE_PI.RES;
    Stoppering_pi.MoveAxis ON FORTE_PI.RES;
    Stoppering_pi.PressStopper ON FORTE_PI.RES;
    Stoppering_pi.RetractPiston ON FORTE_PI.RES;
    Stoppering_pi.Resetting ON FORTE_PI.RES;
    Stoppering_pi.Stopping ON FORTE_PI.RES;
    Stoppering_pi.Stoppering ON FORTE_PI.RES;
  END_MAPPINGS
END_SYSTEM
